Fanuc KAREL source: KD00068.KL

PROGRAM KD00068
%NOLOCKGROUP
VAR
  I: INTEGER
  J: INTEGER
  B: BOOLEAN
  R: REAL
  S: STRING[80]
BEGIN
  CONDITION[1]:
  WHEN DIN[1] = ON DO
    PULSE DOUT[2] FOR 100
  ENDCONDITION
END KD00068
